// TIA Portal V20 export
// export: Created 2026-10-12T16:46:22.9116951Z, ExportSetting WithDefaults, DisplayName Totally Integrated Automation Portal, DisplayVersion V20 Update 6, DisplayName TIA Portal Openness, DisplayVersion V20 Update 6, DisplayName TIA Portal Version Control Interface, DisplayVersion V20 Update 6, DisplayName SINAMICS Startdrive Advanced, DisplayVersion V20 SP1 Update 2, DisplayName SINAMICS Startdrive G110M, G120, G120C, G120D, G120P, G115D, DisplayVersion V20 SP1 Update 2, DisplayName SINAMICS Startdrive G130, G150, S120, S150, SINAMICS MV, G220, S200, S210, DisplayVersion V20 SP1 Update 2, DisplayName STEP 7 Professional, DisplayVersion V20 Update 6, DisplayName STEP 7 Safety, DisplayVersion V20 Update 2, DisplayName WinCC Basic/Comfort/Advanced, DisplayVersion V20 Update 6, DisplayName WinCC Professional, DisplayVersion V20 Update 6, DisplayName WinCC Unified, DisplayVersion V20 Update 6
TYPE "UDT_Prozessroute"
// stored: IsFailsafeCompliant false
   STRUCT
      AuftragsNr : String;
      Kunden : String;
      ID_Artikel : Int;
      ID_Prozessgruppe : Int;
      Personal_ID : Int;
      Anzahl_Schritte : Int;
      Schritte : Array[0..50] of "UDT_Badschritt";
      Freigabe : Bool;
      Abbruch : Bool;
   END_STRUCT;
END_TYPE
